// TIA Portal V21 export
// export: Created 2026-11-10T07:35:25.2706527Z, ExportSetting WithDefaults, DisplayName Totally Integrated Automation Portal, DisplayVersion V21 Update 3, DisplayName STEP 7 Professional, DisplayVersion V21 Update 3, DisplayName STEP 7 Safety, DisplayVersion V21, DisplayName Tech WebApplication, DisplayVersion V21, DisplayName WinCC Basic/Comfort/Advanced, DisplayVersion V21 Update 3, DisplayName WinCC Unified, DisplayVersion V21 Update 3
FUNCTION_BLOCK "FB_Lad_ou004"   // FB76, LAD
{ S7_Optimized_Access := 'TRUE' }
VERSION : 0.1
// stored: AutoNumber true, IsIECCheckEnabled false, IsRetainMemResEnabled false, MemoryReserve 100, SetENOAutomatically false, UDAEnableTagReadback false
   VAR_INPUT
      v_en_r : Bool;
      v_cont : Bool;
      v_len : UDInt;
      v_adhoc : Bool;
   END_VAR
   VAR_OUTPUT
      v_done : Bool;
      v_busy : Bool;
      v_error : Bool;
      v_status : Word;
      v_rcvd_len : UDInt;
   END_VAR
   VAR_IN_OUT
      v_connect : Array[0..99] of Byte;
      v_data : Array[0..99] of Byte;
      v_addr : Array[0..99] of Byte;
      v_com_rst : Bool;
   END_VAR
   VAR
      inst { S7_SetPoint := 'True'} : TRCV_C;
   END_VAR
BEGIN

REGION Network 1: TRCV_C - Establishing a connection and receiving data
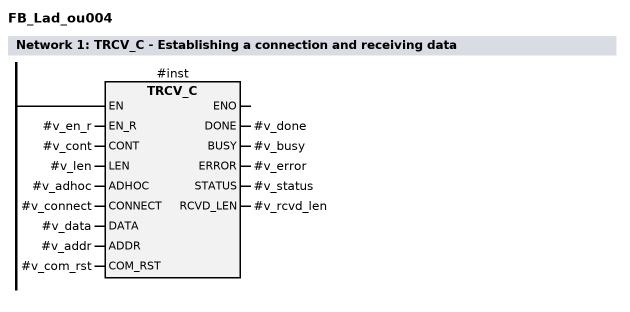
   RUNG wire#powerrail
      #inst.TRCV_C(EN_R := #v_en_r, CONT := #v_cont, LEN := #v_len, ADHOC := #v_adhoc, CONNECT := #v_connect, DATA := #v_data, ADDR := #v_addr, COM_RST := #v_com_rst, DONE => #v_done, BUSY => #v_busy, ERROR => #v_error, STATUS => #v_status, RCVD_LEN => #v_rcvd_len)
   END_RUNG
   // the same network as SCL:
   #inst(EN_R := #v_en_r,   // TRCV_C
         CONT := #v_cont,
         LEN := #v_len,
         ADHOC := #v_adhoc,
         CONNECT := #v_connect,
         DATA := #v_data,
         ADDR := #v_addr,
         COM_RST := #v_com_rst,
         DONE => #v_done,
         BUSY => #v_busy,
         ERROR => #v_error,
         STATUS => #v_status,
         RCVD_LEN => #v_rcvd_len);
END_REGION
END_FUNCTION_BLOCK
